Staubli VAL3: getSize.pgx

public program getSize(num& x_nSize)
begin
  if size(trajTemp:tTrajItem)>0
    x_nSize=size(trajTemp:tTrajItem)
  else
    x_nSize=0
  endIf
end
